{attribute 'qualified_only'}
{attribute 'strict'}
TYPE PlatformKind :
(
	SIMULATION := 0,
	HARDWARE
);
END_TYPE

(* stored: Version 1.1.0.1, ProductVersion 3.1.4026.12
   DUT PlatformKind: Id {118f33c3-84fd-59e8-947b-736266802811} *)
